(* PLC project Vn_return_cond, Beckhoff Automation GmbH TwinCAT PLC Control 3.5.13.21 *)
(* stored: creationDateTime 1970-01-01T00:00:00 *)

PROGRAM Vn_return_cond

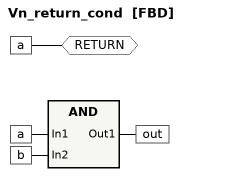
(* FBD diagram, written out as Structured Text *)
IF a THEN RETURN; END_IF;
out := a AND b;
END_PROGRAM
